(* PLC project g_ftrig_edge, Anonymous Benchmark Suite 1.0 *)
(* stored: creationDateTime 2026-07-09T00:00:00 *)

PROGRAM g_ftrig_edge
  VAR_INPUT
    Sig : BOOL;
  END_VAR
  VAR_OUTPUT
    Fall : BOOL;
    OneShot : BOOL;
    Sig_prev : BOOL;
  END_VAR

(* LD diagram, written out as Structured Text *)
Fall := NOT Sig AND Sig_prev;
OneShot := Fall;
Sig_prev := Sig;
END_PROGRAM

CONFIGURATION Config0
  RESOURCE Res0 ON PLC
    TASK tcyclic(INTERVAL := T#10ms, PRIORITY := 0);
    PROGRAM inst0 WITH tcyclic : g_ftrig_edge;
  END_RESOURCE
END_CONFIGURATION
